Fanuc KAREL source: kb00181.KL

PROGRAM KB00181
%STACKSIZE=65535
%PRIORITY=65535
%NOLOCKGROUP
VAR
P1 : INTEGER
BEGIN
P1=1
SET_TIME(P1)
END KB00181
